(* IEC 61131-3 sources: trust-platform/examples/communication/ads_line1/src/generated, 1 file *)

(* ---- ads_generated.st ---- *)
(* Generated by trust-runtime ads import-symbols. Do not edit by hand. *)
TYPE
    ADS_QUALITY : (Stale := 0, Good := 1, Error := 2);
END_TYPE

VAR_GLOBAL
    (* ADS connection: line1 *)
    (* symbol MAIN.Temperature *)
    line1_temp : REAL;
    line1_temp_quality : ADS_QUALITY := Stale;
    (* symbol GVL.LineReady *)
    line1_ready : BOOL;
    line1_ready_quality : ADS_QUALITY := Stale;
    (* symbol GVL.Setpoint *)
    line1_setpoint : REAL;
    line1_setpoint_quality : ADS_QUALITY := Stale;
    (* index group=0x00004020 offset=0x00000000 size=2 *)
    line1_status : WORD;
    line1_status_quality : ADS_QUALITY := Stale;
END_VAR
